// TIA Portal V20 export
TYPE "WT3_Plattform_Status_UDT"
   STRUCT
      iHandshake : Int;
      Datum : Array[0..9] of Char;
      Zeit : Array[0..7] of Char;
      SwVersion : Array[0..7] of Char;
      Alarm : Struct
         bE0000_KonfigAlarm : Bool;
         bE0001_IOZuweisungUnvollst : Bool;
         bE0002_Reserviert : Bool;
         bE0003_Reserviert : Bool;
         bE0004_AlarmIOKomm : Bool;
         bE0005_AlarmKabelbruch : Bool;
         bE0006_AlarmIOHWKonfig : Bool;
         bE0007_Reserviert : Bool;
         bE0008_Reserviert : Bool;
         bE0009_Reserviert : Bool;
         bE0010_Reserviert : Bool;
         bE0011_Reserviert : Bool;
         bE0012_Reserviert : Bool;
         bE0013_Reserviert : Bool;
         bE0014_Reserviert : Bool;
         bE0015_Reserviert : Bool;
         bE0016_Reserviert : Bool;
         bE0017_AlarmKeineLizenzVorhanden : Bool;
         b302_Reserve : Bool;
         b303_Reserve : Bool;
         b304_Reserve : Bool;
         b305_Reserve : Bool;
         b306_Reserve : Bool;
         b307_Reserve : Bool;
         by31_Reserve : Byte;
         by32_Reserve : Byte;
         by33_Reserve : Byte;
         by34_Reserve : Byte;
         by35_Reserve : Byte;
         by36_Reserve : Byte;
         by37_Reserve : Byte;
         by38_Reserve : Byte;
         by39_Reserve : Byte;
         by40_Reserve : Byte;
         by41_Reserve : Byte;
         by42_Reserve : Byte;
         by43_Reserve : Byte;
         by44_Reserve : Byte;
         by45_Reserve : Byte;
         by46_Reserve : Byte;
         by47_Reserve : Byte;
         by48_Reserve : Byte;
         by49_Reserve : Byte;
         by50_Reserve : Byte;
         by51_Reserve : Byte;
         by52_Reserve : Byte;
         by53_Reserve : Byte;
         by54_Reserve : Byte;
         by55_Reserve : Byte;
         by56_Reserve : Byte;
         by57_Reserve : Byte;
         by58_Reserve : Byte;
         by59_Reserve : Byte;
      END_STRUCT;
      Warnung : Struct
         bA1000_Reserviert : Bool;
         bA1001_Reserviert : Bool;
         bA1002_Reserviert : Bool;
         bA1003_Reserviert : Bool;
         bA1004_Reserviert : Bool;
         bA1005_WarnungKabelbruch : Bool;
         bA1006_Reserviert : Bool;
         bA1007_WarnungFeldbus : Bool;
         bA1008_Reserviert : Bool;
         bA1009_Reserviert : Bool;
         bA1010_WarnungbeiInitialisierungSteuerkommunikation : Bool;
         bA1011_Reserviert : Bool;
         bA1012_Reserviert : Bool;
         bA1013_Reserviert : Bool;
         bA1014_Reserviert : Bool;
         bA1015_Reserviert : Bool;
         bA1016_Reserviert : Bool;
         bA1017_WarnungKeineLizenzVorhanden : Bool;
         bA1018_WarnungSpeisungHeizung230V : Bool;
         bA1019_WarnungSelektivitätsmodul : Bool;
         bA1020_WarnungLastschalter : Bool;
         bA1021_WarnungHauptschalter : Bool;
         bA1022_WarnungHauptkontakteLaststromkreis : Bool;
         "bA1023_WarnungI/O-KommunikationWT3" : Bool;
         "bA1024_WarnungI/O-KonfigurationWT3" : Bool;
         b631_Reserve : Bool;
         b632_Reserve : Bool;
         b633_Reserve : Bool;
         b634_Reserve : Bool;
         b635_Reserve : Bool;
         b636_Reserve : Bool;
         b637_Reserve : Bool;
         by64_Reserve : Byte;
         by65_Reserve : Byte;
         by66_Reserve : Byte;
         by67_Reserve : Byte;
         by68_Reserve : Byte;
         by69_Reserve : Byte;
         by70_Reserve : Byte;
         by71_Reserve : Byte;
         by72_Reserve : Byte;
         by73_Reserve : Byte;
         by74_Reserve : Byte;
         by75_Reserve : Byte;
         by76_Reserve : Byte;
         by77_Reserve : Byte;
         by78_Reserve : Byte;
         by79_Reserve : Byte;
         by80_Reserve : Byte;
         by81_Reserve : Byte;
         by82_Reserve : Byte;
         by83_Reserve : Byte;
         by84_Reserve : Byte;
         by85_Reserve : Byte;
         by86_Reserve : Byte;
         by87_Reserve : Byte;
         by88_Reserve : Byte;
         by89_Reserve : Byte;
         by90_Reserve : Byte;
         by91_Reserve : Byte;
      END_STRUCT;
      Zustand : Struct
         bAlarmzustandAktiv : Bool;
         bWarnzustandAktiv : Bool;
         bSystemMeldungAktiv : Bool;
         bSeviceMeldungAktiv : Bool;
         bStopManuell : Bool;
         bStopAuto : Bool;
         bStopExtern : Bool;
         bBetriebAuto : Bool;
         bBetriebManuell : Bool;
         bAnlaufAuto : Bool;
         bAnlaufManuell : Bool;
         bManuellStoppen : Bool;
         b934_Reserve : Bool;
         b935_Reserve : Bool;
         b936_Reserve : Bool;
         b937_Reserve : Bool;
         by94_Reserve : Byte;
         bSystemMeldungKonfigUmschaltung : Bool;
         b951_Reserve : Bool;
         b952_Reserve : Bool;
         b953_Reserve : Bool;
         b954_Reserve : Bool;
         b955_Reserve : Bool;
         b956_Reserve : Bool;
         b957_Reserve : Bool;
         by96_Reserve : Byte;
         by97_Reserve : Byte;
         by98_Reserve : Byte;
         by99_Reserve : Byte;
         by100_Reserve : Byte;
         by101_Reserve : Byte;
         by102_Reserve : Byte;
         by103_Reserve : Byte;
         by104_Reserve : Byte;
         by105_Reserve : Byte;
         by106_Reserve : Byte;
         by107_Reserve : Byte;
      END_STRUCT;
      DigIn : Struct
         bKonfigSatzBit0 : Bool;
         bKonfigSatzBit1 : Bool;
         bFreigabeTempRegler : Bool;
         bFreigabeZweipunktRegler1 : Bool;
         bFreigabeZweipunktRegler2 : Bool;
         bFreigabeZweipunktregler3 : Bool;
         bFreigabeZweipunktregler4 : Bool;
         bFreigabePIRegler1 : Bool;
         bFreigabePIRegler2 : Bool;
         bFreigabePIRegler3 : Bool;
         bFreigabePIRegler4 : Bool;
         bPiRegler1SollwertB : Bool;
         bPiRegler2SollwertB : Bool;
         bPiRegler3SollwertB : Bool;
         bPiRegler4SollwertB : Bool;
         bAuxDigital1 : Bool;
         bAuxDigital2 : Bool;
         bAuxDigital3 : Bool;
         bAuxDigital4 : Bool;
         bAuxDigital5 : Bool;
         bAuxDigital6 : Bool;
         bAuxDigital7 : Bool;
         bAuxDigital8 : Bool;
         b1107_Reserve : Bool;
         by111_Reserve : Byte;
         by112_Reserve : Byte;
         by113_Reserve : Byte;
         by114_Reserve : Byte;
         by115_Reserve : Byte;
      END_STRUCT;
      DigOut : Struct
         bAlarm : Bool;
         bWarnung : Bool;
         bTemperaturregler : Bool;
         bZweipunktrelger1 : Bool;
         bZweipunktrelger2 : Bool;
         bZweipunktregler3 : Bool;
         bZweipunktregler4 : Bool;
         bQDigitaleVerknüpfung1 : Bool;
         bQDigitaleVerknüpfung2 : Bool;
         bQDigitaleVerknüpfung3 : Bool;
         bQDigitaleVerknüpfung4 : Bool;
         bQDigitaleVerknüpfung5 : Bool;
         bQDigitaleVerknüpfung6 : Bool;
         bQDigitaleVerknüpfung7 : Bool;
         bQDigitaleVerknüpfung8 : Bool;
         bQDigitaleVerknüpfung9 : Bool;
         bQDigitaleVerknüpfung10 : Bool;
         bQDigitaleVerknüpfung11 : Bool;
         bQDigitaleVerknüpfung12 : Bool;
         bQInverter1 : Bool;
         bQInverter2 : Bool;
         bQInverter3 : Bool;
         bQInverter4 : Bool;
         bQZeitglied1 : Bool;
         bQZeitglied2 : Bool;
         bQZeitglied3 : Bool;
         bQZeitglied4 : Bool;
         bQRsFlipFlop1 : Bool;
         bQRsFlipFlop2 : Bool;
         bQRsFlipFlop3 : Bool;
         bQRsFlipFlop4 : Bool;
         bQRsFlipFlop5 : Bool;
         bQRsFlipFlop6 : Bool;
         bQRsFlipFlop7 : Bool;
         bQRsFlipFlop8 : Bool;
         bQRsFlipFlop9 : Bool;
         bQRsFlipFlop10 : Bool;
         bQRsFlipFlop11 : Bool;
         bQRsFlipFlop12 : Bool;
         bQDigitaleVerknüpfung13 : Bool;
         bQDigitaleVerknüpfung14 : Bool;
         bQDigitaleVerknüpfung15 : Bool;
         bQDigitaleVerknüpfung16 : Bool;
         bSammelkanal1 : Bool;
         bSammelkanal2 : Bool;
         bSammelkanal3 : Bool;
         bSammelkanal4 : Bool;
         bSammelkanal5 : Bool;
         bSammelkanal6 : Bool;
         b1221_Reserve : Bool;
         b1222_Reserve : Bool;
         b1223_Reserve : Bool;
         b1224_Reserve : Bool;
         b1225_Reserve : Bool;
         b1226_Reserve : Bool;
         b1227_Reserve : Bool;
         by123_Reserve : Byte;
      END_STRUCT;
      iKonfigSatz : Int;
      rZweipunktregler1Istwert : Real;
      rZweipunktregler2Istwert : Real;
      rZweipunktregler3Istwert : Real;
      rZweipunktregler4Istwert : Real;
      rPiRegler1Istwert : Real;
      rPiRegler1Sollwert : Real;
      diPiRegler1Sollwertrampe : DInt;
      rPiRegler1Stellwert : Real;
      rPiRegler2Istwert : Real;
      rPiRegler2Sollwert : Real;
      diPiRegler2Sollwertrampe : DInt;
      rPiRegler2Stellwert : Real;
      rPiRegler3Istwert : Real;
      rPiRegler3Sollwert : Real;
      diPiRegler3Sollwertrampe : DInt;
      rPiRegler3Stellwert : Real;
      rPiRegler4Istwert : Real;
      rPiRegler4Sollwert : Real;
      diPiRegler4Sollwertrampe : DInt;
      rPiRegler4Stellwert : Real;
      rI1AnalogeVerknüpfung1 : Real;
      rI2AnalogeVerknüpfung1 : Real;
      rQAnalogeVerknüpfung1 : Real;
      rI1AnalogeVerknüpfung2 : Real;
      rI2AnalogeVerknüpfung2 : Real;
      rQAnalogeVerknüpfung2 : Real;
      rI1AnalogeVerknüpfung3 : Real;
      rI2AnalogeVerknüpfung3 : Real;
      rQAnalogeVerknüpfung3 : Real;
      rI1AnalogeVerknüpfung4 : Real;
      rI2AnalogeVerknüpfung4 : Real;
      rQAnalogeVerknüpfung4 : Real;
      rI1AnalogeVerknüpfung5 : Real;
      rI2AnalogeVerknüpfung5 : Real;
      rQAnalogeVerknüpfung5 : Real;
      rI1AnalogeVerknüpfung6 : Real;
      rI2AnalogeVerknüpfung6 : Real;
      rQAnalogeVerknüpfung6 : Real;
      rI1AnalogeVerknüpfung7 : Real;
      rI2AnalogeVerknüpfung7 : Real;
      rQAnalogeVerknüpfung7 : Real;
      rI1AnalogeVerknüpfung8 : Real;
      rI2AnalogeVerknüpfung8 : Real;
      rQAnalogeVerknüpfung8 : Real;
      rI1AnalogeVerknüpfung9 : Real;
      rI2AnalogeVerknüpfung9 : Real;
      rQAnalogeVerknüpfung9 : Real;
      rI1AnalogeVerknüpfung10 : Real;
      rI2AnalogeVerknüpfung10 : Real;
      rQAnalogeVerknüpfung10 : Real;
      rI1AnalogeVerknüpfung11 : Real;
      rI2AnalogeVerknüpfung11 : Real;
      rQAnalogeVerknüpfung11 : Real;
      rI1AnalogeVerknüpfung12 : Real;
      rI2AnalogeVerknüpfung12 : Real;
      rQAnalogeVerknüpfung12 : Real;
      rISequenz1 : Real;
      rQSequenz1 : Real;
      rISequenz2 : Real;
      rQSequenz2 : Real;
      rISequenz3 : Real;
      rQSequenz3 : Real;
      rISequenz4 : Real;
      rQSequenz4 : Real;
      rISequenz5 : Real;
      rQSequenz5 : Real;
      rISequenz6 : Real;
      rQSequenz6 : Real;
      rISequenz7 : Real;
      rQSequenz7 : Real;
      rISequenz8 : Real;
      rQSequenz8 : Real;
      rISequenz9 : Real;
      rQSequenz9 : Real;
      rISequenz10 : Real;
      rQSequenz10 : Real;
      rISequenz11 : Real;
      rQSequenz11 : Real;
      rISequenz12 : Real;
      rQSequenz12 : Real;
      rIUmrechnung1 : Real;
      rQUmrechnung1 : Real;
      rIUmrechnung2 : Real;
      rQUmrechnung2 : Real;
      rIUmrechnung3 : Real;
      rQUmrechnung3 : Real;
      rIUmrechnung4 : Real;
      rQUmrechnung4 : Real;
      rIRampe1 : Real;
      rQRampe1 : Real;
      rIRampe2 : Real;
      rQRampe2 : Real;
      rIRampe3 : Real;
      rQRampe3 : Real;
      rIRampe4 : Real;
      rQRampe4 : Real;
      byReserve : Array[510..629] of Byte;
   END_STRUCT;
END_TYPE
